(* IEC 61131-3 sources: plcassist-cli/packages/volt-lsp-iec/test-corpus/awa-palletizer/Device/Plc Logic/Application/Library Manager/SysCpuHandling, 11 files *)

(* ---- SYSCPUATOMICADD.fun ---- *)
FUNCTION SYSCPUATOMICADD : DINT
VAR_INPUT
	PIVALUE : POINTER TO DINT;
	NSUM : DINT;
	PRESULT : POINTER TO RTS_IEC_RESULT;
END_VAR
END_FUNCTION

(* ---- SYSCPUATOMICADD64.fun ---- *)
FUNCTION SYSCPUATOMICADD64 : LINT
VAR_INPUT
	PIVALUE : POINTER TO LINT;
	NSUM : LINT;
	PRESULT : POINTER TO RTS_IEC_RESULT;
END_VAR
END_FUNCTION

(* ---- SYSCPUATOMICCOMPAREANDSWAP.fun ---- *)
FUNCTION SYSCPUATOMICCOMPAREANDSWAP : RTS_IEC_RESULT
VAR_INPUT
	PADDRESS : POINTER TO BYTE;
	PSWAPVALUE : POINTER TO BYTE;
	PCOMPAREVALUE : POINTER TO BYTE;
	VALUESIZE : USINT;
END_VAR
END_FUNCTION

(* ---- SYSCPUCALLIECFUNCWITHPARAMS.fun ---- *)
FUNCTION SYSCPUCALLIECFUNCWITHPARAMS : RTS_IEC_RESULT
VAR_INPUT
	PFIECFUNC : POINTER TO BYTE;
	PPARAM : POINTER TO BYTE;
	ULSIZE : UDINT;
END_VAR
END_FUNCTION

(* ---- SYSCPURESETBIT.fun ---- *)
FUNCTION SYSCPURESETBIT : RTS_IEC_RESULT
VAR_INPUT
	PULVALUE : POINTER TO UDINT;
	ULBIT : UDINT;
END_VAR
END_FUNCTION

(* ---- SYSCPURESETBIT2.fun ---- *)
FUNCTION SYSCPURESETBIT2 : RTS_IEC_RESULT
VAR_INPUT
	PBYVALUE : POINTER TO BYTE;
	ULBIT : UDINT;
END_VAR
END_FUNCTION

(* ---- SYSCPUSETBIT.fun ---- *)
FUNCTION SYSCPUSETBIT : RTS_IEC_RESULT
VAR_INPUT
	PULVALUE : POINTER TO UDINT;
	ULBIT : UDINT;
END_VAR
END_FUNCTION

(* ---- SYSCPUSETBIT2.fun ---- *)
FUNCTION SYSCPUSETBIT2 : RTS_IEC_RESULT
VAR_INPUT
	PBYVALUE : POINTER TO BYTE;
	ULBIT : UDINT;
END_VAR
END_FUNCTION

(* ---- SYSCPUTESTANDRESET.fun ---- *)
FUNCTION SYSCPUTESTANDRESET : RTS_IEC_RESULT
VAR_INPUT
	PULVALUE : POINTER TO UDINT;
	ULBIT : UDINT;
END_VAR
END_FUNCTION

(* ---- SYSCPUTESTANDSET.fun ---- *)
FUNCTION SYSCPUTESTANDSET : RTS_IEC_RESULT
VAR_INPUT
	PULVALUE : POINTER TO UDINT;
	ULBIT : UDINT;
END_VAR
END_FUNCTION

(* ---- SYSCPUTESTANDSETBIT.fun ---- *)
FUNCTION SYSCPUTESTANDSETBIT : RTS_IEC_RESULT
VAR_INPUT
	PADDRESS : POINTER TO BYTE;
	NLEN : UDINT;
	IBIT : DINT;
	BSET : DINT;
END_VAR
END_FUNCTION
